// TIA Portal V19 export
// export: Created 2026-10-15T10:10:37.3882165Z, ExportSetting WithDefaults, DisplayName Totally Integrated Automation Portal, DisplayVersion V19, DisplayName TIA Portal Openness, DisplayVersion V19, DisplayName TIA Portal Version Control Interface, DisplayVersion V19, DisplayName STEP 7 Professional, DisplayVersion V19, DisplayName STEP 7 Safety, DisplayVersion V19, DisplayName WinCC Basic/Comfort/Advanced, DisplayVersion V19, DisplayName WinCC Unified, DisplayVersion V19
FUNCTION "ROLL_Cycle" : Void   // FC39, SCL
{ S7_Optimized_Access := 'TRUE' }
VERSION : 0.1
// stored: AutoNumber true, IsIECCheckEnabled false, SetENOAutomatically false, UDAEnableTagReadback false
   VAR_TEMP
      delta : LReal;
   END_VAR
BEGIN

   #delta := RUNTIME("ROLL_IO".RuntimeMemory) * 1000.0;
   IF "ROLL_IO".FirstCycle THEN
       #delta := 0.0;
       "ROLL_IO".FirstCycle := FALSE;
   END_IF;
   "ROLL_ReadInputs"();
   "ROLL_AdvanceTime"(DeltaMs := #delta);
   // Exact OB1 order for the process blocks; startup DB creation is replaced.
   IF NOT "ROLL_State".M[0, 2] THEN
       "ROLL_State".M[0, 1] := FALSE;
   END_IF;
   IF "ROLL_State".M[0, 1] THEN
       "ROLL_State".M[0, 7] := TRUE;
   END_IF;
   "ROLL_State".M[0, 5] := NOT "ROLL_State".M[0, 5];
   IF "ROLL_State".M[3, 2] THEN
       "ROLL_State".M[3, 3] := TRUE;
   END_IF;
   IF "ROLL_IO".Input[0, 2] THEN
       "ROLL_State".M[3, 3] := FALSE;
   END_IF;
   "ROLL_State".M[3, 2] := "ROLL_IO".Input[0, 1] AND NOT "ROLL_State".M[0, 1];
   "ROLL_PB2"();
   IF "ROLL_State".M[0, 7] THEN
       "ROLL_State".M[0, 7] := FALSE;
   END_IF;
   "ROLL_PB3"();
   "ROLL_PB4"();
   "ROLL_PB19"();
   "ROLL_PB21"();
   "ROLL_PB50"();
   "ROLL_PB51"();
   "ROLL_PB52"();
   IF NOT "ROLL_State".M[3, 3] THEN
       "ROLL_PB8"();
   END_IF;
   IF NOT "ROLL_State".M[3, 3] THEN
       "ROLL_PB9"();
   END_IF;
   IF NOT "ROLL_State".M[3, 3] THEN
       "ROLL_PB10"();
   END_IF;
   IF NOT "ROLL_State".M[3, 3] THEN
       "ROLL_PB14"();
   END_IF;
   IF "ROLL_State".M[3, 3] THEN
       "ROLL_PB16"();
   END_IF;
   "ROLL_PB7"();
   "ROLL_PB13"();
   "ROLL_PB15"();
   "ROLL_PB17"();
   "ROLL_PB20"();
   "ROLL_PB23"();
   "ROLL_PB24"();
   "ROLL_PB25"();
   "ROLL_FB111"();
   "ROLL_HmiExchange"(DeltaMs := #delta);
   "ROLL_WriteOutputs"();
END_FUNCTION
